FUNCTION_BLOCK CAN_MSG_TO_STRING (* CAN_MSG von AlPgnRxNew8B (bis 8 Byte) als STRING auslesen *)
  (* Standard: 61499-2; Description: Copyright (c) 2026 HR Agrartechnik GmbH This program and the accompanying materials are made available under the terms of the Eclipse Public License 2.0 which is available at https://www.eclipse.org/legal/epl-2.0/ SPDX-License-Identifier: EPL-2.0 *)
  (* Version 1.1, 2026-11-14, Franz Höpfinger, HR Agrartechnik GmbH, unnoetige Konvertierungen UINT_TO_DINT/CHAR_TO_STRING entfernt (IDE-Warnungen) *)
  (* Version 1.0, 2026-11-13, Franz Höpfinger, HR Agrartechnik GmbH, Initial Version - STRING ueber CAN (0-8 Byte) *)
  PACKAGE isobus::pgn;
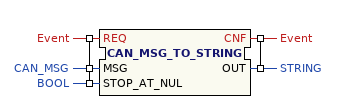
  EVENT_INPUT
    REQ WITH MSG, STOP_AT_NUL; (* Text auslesen *)
  END_EVENT
  EVENT_OUTPUT
    CNF WITH OUT; (* OUT ist gefuellt *)
  END_EVENT
  VAR_INPUT
    MSG : isobus::pgn::CAN_MSG; (* empfangene Nachricht, gelesen werden u16DaSize Bytes (hoechstens 8) *)
    STOP_AT_NUL : BOOL := TRUE; (* TRUE: Text endet vor dem ersten 16#00 *)
  END_VAR
  VAR_OUTPUT
    OUT : STRING; (* Text, je Byte 1 Zeichen *)
  END_VAR
  EC_STATES
    REQ : REQ -> CNF;
  END_STATES
  ALGORITHM REQ IN ST: (* data[0..u16DaSize-1] als Zeichen anhaengen *)
VAR_TEMP
	n : DINT; // Anzahl zu lesender Bytes
	i : DINT; // Laufindex
	b : BYTE; // aktuelles Byte
END_VAR
OUT := '';
n := MSG.u16DaSize;
IF n > 8 THEN
	n := 8;
END_IF;
FOR i := 1 TO n DO
	b := MSG.data[i - 1];
	IF STOP_AT_NUL AND (b = BYTE#0) THEN
		EXIT;
	END_IF;
	OUT := CONCAT(OUT, BYTE_TO_CHAR(b));
END_FOR;
  END_ALGORITHM
END_FUNCTION_BLOCK
